FUNCTION_BLOCK MUX_MY (* Basic Function Block Type *)
  (* Standard: 61499-2 *)
  (* Version 0.0, 10/19/2026, macie, Schneider Electric, Template *)
  PACKAGE Main;
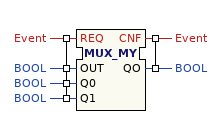
  EVENT_INPUT
    REQ WITH OUT, Q0, Q1; (* Normal Execution Request *)
  END_EVENT
  EVENT_OUTPUT
    CNF WITH QO; (* Execution Confirmation *)
  END_EVENT
  VAR_INPUT
    OUT : BOOL;
    Q0 : BOOL; (* Input event qualifier *)
    Q1 : BOOL;
  END_VAR
  VAR_OUTPUT
    QO : BOOL; (* Output event qualifier *)
  END_VAR
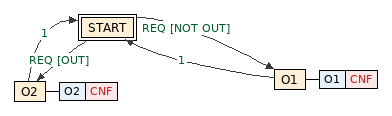
  EC_STATES
    START; (* Initial State *)
    O2 : O2 -> CNF; (* Normal execution *)
    O1 : O1 -> CNF;
  END_STATES
  EC_TRANSITIONS
    START TO O2 := REQ [OUT];
    O2 TO START := 1;
    START TO O1 := REQ [NOT OUT];
    O1 TO START := 1;
  END_TRANSITIONS
  ALGORITHM O2 IN ST: (* Normally executed algorithm *)
;
QO := Q1;
  END_ALGORITHM
  ALGORITHM O1 IN ST:
;
QO := Q0;
  END_ALGORITHM
END_FUNCTION_BLOCK
